Yaskawa INFORM job: TEAM2V2.JBI

/JOB
//NAME TEAM2V2
//POS
///NPOS 19,0,19,0,0,0
///TOOL 0
///POSTYPE PULSE
///PULSE
C00000=-947,-55524,-59539,-219,-89999,0
C00001=-14550,47390,-9918,-1666,-46835,4504
C00002=-14208,46659,-14977,-1765,-43895,4451
C00003=-14208,46659,-14977,-1765,-43895,4451
C00004=-12937,47080,-14663,-1785,-43777,4060
C00005=2104,31679,-43283,25276,-25005,12090
C00006=-2259,20876,-60136,2215,-15221,39909
C00007=21917,8400,-41377,7972,-38642,30634
C00008=1813,-26553,-79210,-1109,-5821,4862
C00009=1813,-26553,-79210,-1109,-5821,4862
C00010=-13828,10438,-65699,5058,-1053,2039
C00011=-14008,16266,-68247,1762,5093,3588
C00012=-13949,16746,-68323,1395,5510,3745
C00013=-20003,17976,-66586,25043,5725,-5712
C00014=-22190,3498,-80684,50309,12417,-18076
C00015=-23949,17256,-92201,19409,43880,-2545
C00016=-25442,14078,-97059,20257,44843,-2451
C00017=-25442,-290,-95405,25953,33870,-5925
C00018=-947,-55524,-59539,-219,-89999,0
EC00000=-1645
EC00001=-1645
EC00002=-1645
EC00003=-1645
EC00004=-1645
EC00005=-1645
EC00006=-1645
EC00007=-1645
EC00008=-1644
EC00009=-83284
EC00010=-83284
EC00011=-83284
EC00012=-83284
EC00013=-83284
EC00014=-162295
EC00015=-162295
EC00016=-162295
EC00017=-162295
EC00018=-1645
//INST
///DATE 2025/10/20 18:25
///ATTR SC,RW
///GROUP1 RB1,ST1
NOP
MOVJ C00000 EC00000 VJ=0.78
MOVJ C00001 EC00001 VJ=0.78
MOVL C00002 EC00002 V=11.0
ARCON ASF#(65)
MOVC C00003 EC00003 V=11.0
MOVC C00004 EC00004 V=11.0
MOVC C00005 EC00005 V=11.0
MOVC C00006 EC00006 V=11.0
MOVJ C00007 EC00007 VJ=0.78
MOVS C00008 EC00008 V=11.0
MOVS C00009 EC00009 V=11.0
MOVJ C00010 EC00010 VJ=0.78
MOVL C00011 EC00011 V=11.0
ARCON ASF#(65)
MOVL C00012 EC00012 V=11.0
MOVL C00013 EC00013 V=11.0
ARCOF AEF#(65)
MOVJ C00014 EC00014 VJ=0.78
MOVL C00015 EC00015 V=11.0
ARCON ASF#(65)
MOVL C00016 EC00016 V=11.0
ARCOF AEF#(65)
MOVL C00017 EC00017 V=11.0
MOVL C00018 EC00018 V=11.0
END
